Staubli VAL3: trajTemp.dtx

public trajItem tTrajItem{}
